Staubli VAL3: goSafeHome.dtx

mdesc mHome = {accel=25, vel=50, decel=25, blend=off}
mdesc mNomSpeed
